  rq_init_comm_if_connected(9, "1")
  rq_init_comm_if_connected(2, "2")
  rq_init_comm_if_connected(3, "3")
  rq_init_comm_if_connected(4, "4")
  rq_print_connected_grippers()
  rq_gripper_communication_thread = run rq_gripper_communication()
  set_closed_norm(97.6470588235294, "1")
  set_open_norm(1.1764705882352942, "1")
  set_closed_mm(0.0, "1")
  set_open_mm(53.0, "1")
  set_closed_norm(100.0, "2")
  set_open_norm(0.0, "2")
  set_closed_mm(0.0, "2")
  set_open_mm(50.0, "2")
  set_closed_norm(100.0, "3")
  set_open_norm(0.0, "3")
  set_closed_mm(0.0, "3")
  set_open_mm(50.0, "3")
  set_closed_norm(100.0, "4")
  set_open_norm(0.0, "4")
  set_closed_mm(0.0, "4")
  set_open_mm(50.0, "4")
  rq_current_limit_enabled = False
  while(not rq_gripper_communication_thread_started):
      sleep(0.008)
  end
  # end: URCap Installation Node
  step_count_652fcfe5_f3e5_4323_a28e_c4dd7c99f65c = 0.0
  thread Step_Counter_Thread_2d5c0d0e_2884_4a5b_ab92_48b0595c18f1():
    while (True):
      step_count_652fcfe5_f3e5_4323_a28e_c4dd7c99f65c = step_count_652fcfe5_f3e5_4323_a28e_c4dd7c99f65c + 1.0
      sync()
    end
  end
  run Step_Counter_Thread_2d5c0d0e_2884_4a5b_ab92_48b0595c18f1()
  global AMR_Position=struct(position_identifier=0, x1=0, x2=0, y1=0, y2=0, theta1=0, theta2=0)
  $ 2 "BeforeStart"
  $ 3 "Manual"
  $ 4 "Home (Safe)"
  movej([-1.2291867130198177, -1.2978880085432127, -1.8023901537060905, -1.6126269993759976, 1.5736085024106596, 0.3398721000491988], a=1.3962634015954636, v=1.0471975511965976)
  $ 5 "STATE≔'state'"
  global STATE=request_integer_from_primary_client("state")
  $ 6 "If STATE≟6"
  if (STATE == 6):
    $ 7 "Action≔'what'"
    global Action=request_integer_from_primary_client("what")
    $ 8 "If Action≟52"
    if (Action == 52):
      $ 9 "AMR_PosTarget≔'target'"
      global AMR_PosTarget=request_integer_from_primary_client("target")
    end
  end
  $ 10 "Robot Program"
  $ 11 "PreSettings"
  $ 12 "AMR_TargetList≔[1,2,3,4,5,21,22,23,24,31,32,33,34,35,36,37,38,41]"
  global AMR_TargetList=[1,2,3,4,5,21,22,23,24,31,32,33,34,35,36,37,38,41]
  $ 13 "AMR_Done≔ False "
  global AMR_Done=  False
  $ 14 "AMR_PosActual≔T2O_Current_Pos"
  global AMR_PosActual=modbus_get_signal_status("T2O_Current_Pos")
  $ 15 "AMR_Attemps≔T2O_Nav_Attemps"
  global AMR_Attemps=modbus_get_signal_status("T2O_Nav_Attemps")
  $ 16 "AMR_Battery≔MiR_Battery_Lvl"
  global AMR_Battery=modbus_get_signal_status("MiR_Battery_Lvl")
  $ 17 "AMR_Charging≔(T2O_Charging≟1)"
  global AMR_Charging=(modbus_get_signal_status("T2O_Charging") == 1)
  $ 18 "AMR_Position≔struct(position_identifier=T2O_Current_Pos, x1=MiR_Position_X1, x2=MiR_Position_X2, y1=MiR_Position_Y1, y2=MiR_Position_Y2, theta1=MiR_Theta_1, theta2=MiR_Theta_2) "
  global AMR_Position=struct(position_identifier=modbus_get_signal_status("T2O_Current_Pos"), x1=modbus_get_signal_status("MiR_Position_X1"), x2=modbus_get_signal_status("MiR_Position_X2"), y1=modbus_get_signal_status("MiR_Position_Y1"), y2=modbus_get_signal_status("MiR_Position_Y2"), theta1=modbus_get_signal_status("MiR_Theta_1"), theta2=modbus_get_signal_status("MiR_Theta_2"))
  $ 19 "If MiR_Mode≠7"
  if (modbus_get_signal_status("MiR_Mode") != 7):
    $ 20 "Error"
    $ 21 "set_error(ERROR_AMR_WRONG_MODE)"
    set_error(ERROR_AMR_WRONG_MODE)
    $ 22 "AMR_Done≔ True "
    global AMR_Done=  True
  end
  $ 23 "'=========='"
  # '=========='
  $ 24 "Switch STATE"
  switch_1 = STATE
  $ 25 "Case 1"
  if (1 == switch_1):
    $ 26 "stopping"
    $ 27 "If T2O_Done≟1 and O2T_Acknowledge≟0"
    if (modbus_get_signal_status("T2O_Done") == 1  and  modbus_get_signal_status("O2T_Acknowledge") == 0):
      $ 28 "Set O2T_Acknowledge=1"
      modbus_set_output_register("O2T_Acknowledge", 1)
    end
    $ 29 "Set MiR_CMD_Stop=On"
    modbus_set_output_signal("MiR_CMD_Stop", True)
    $ 30 "If MiR_State≠3 and MiR_State≠5"
    if (modbus_get_signal_status("MiR_State") != 3  and  modbus_get_signal_status("MiR_State") != 5):
      $ 31 "AMR_Position.position_identifier = 0"
      AMR_Position.position_identifier = 0
      $ 32 "AMR_Done≔ True "
      global AMR_Done=  True
    end
  elif (2 == switch_1):
    $ 33 "Case 2"
    $ 34 "stopped"
    $ 35 "Set MiR_CMD_Stop=Off"
    modbus_set_output_signal("MiR_CMD_Stop", False)
  elif (3 == switch_1):
    $ 36 "Case 3"
    $ 37 "resetting"
    $ 38 "Set O2T_Mis_Main=Off"
    modbus_set_output_signal("O2T_Mis_Main", False)
    $ 39 "Set O2T_Mis_Charge=Off"
    modbus_set_output_signal("O2T_Mis_Charge", False)
    $ 40 "If MiR_Mis_Queue>0"
    if (modbus_get_signal_status("MiR_Mis_Queue")>0):
      $ 41 "Set MiR_CMD_Clear_Q=On"
      modbus_set_output_signal("MiR_CMD_Clear_Q", True)
      $ 42 "Wait MiR_Mis_Queue≟0"
      while (not(modbus_get_signal_status("MiR_Mis_Queue") == 0)):
        sync()
      end
      $ 43 "Set MiR_CMD_Clear_Q=Off"
      modbus_set_output_signal("MiR_CMD_Clear_Q", False)
    end
    $ 44 "If MiR_Error_ID≠0"
    if (modbus_get_signal_status("MiR_Error_ID") != 0):
      $ 45 "Set MiR_CMD_Clear_E=On"
      modbus_set_output_signal("MiR_CMD_Clear_E", True)
      $ 46 "Wait MiR_Error_ID≟0"
      while (not(modbus_get_signal_status("MiR_Error_ID") == 0)):
        sync()
      end
      $ 47 "Set MiR_CMD_Clear_E=Off"
      modbus_set_output_signal("MiR_CMD_Clear_E", False)
    end
    $ 48 "Set O2T_Action=0"
    modbus_set_output_register("O2T_Action", 0)
    $ 49 "Set O2T_Acknowledge=0"
    modbus_set_output_register("O2T_Acknowledge", 0)
    $ 50 "Set O2T_Target_Pos=0"
    modbus_set_output_register("O2T_Target_Pos", 0)
    $ 51 "Set O2T_Footprint=0"
    modbus_set_output_register("O2T_Footprint", 0)
    $ 52 "Set O2T_ProtectOff=0"
    modbus_set_output_register("O2T_ProtectOff", 0)
    $ 53 "Set O2T_Dock=0"
    modbus_set_output_register("O2T_Dock", 0)
    $ 54 "AMR_Attemps≔0"
    global AMR_Attemps=0
    $ 55 "AMR_PosTarget≔0"
    global AMR_PosTarget=0
    $ 56 "AMR_Step≔0"
    global AMR_Step=0
    $ 57 "AMR_AtTarget≔ False "
    global AMR_AtTarget=  False
    $ 58 "If MiR_State≟4 or MiR_State≟3 or MiR_State≟10"
    if (modbus_get_signal_status("MiR_State") == 4  or  modbus_get_signal_status("MiR_State") == 3  or  modbus_get_signal_status("MiR_State") == 10):
      $ 59 "AMR_Done≔ True "
      global AMR_Done=  True
    end
  elif (5 == switch_1):
    $ 60 "Case 5"
    $ 61 "starting"
    $ 62 "If MiR_State≟4"
    if (modbus_get_signal_status("MiR_State") == 4):
      $ 63 "Set MiR_CMD_Start=On"
      modbus_set_output_signal("MiR_CMD_Start", True)
      $ 64 "Wait MiR_State≠4"
      while (not(modbus_get_signal_status("MiR_State") != 4)):
        sync()
      end
      $ 65 "Set MiR_CMD_Start=Off"
      modbus_set_output_signal("MiR_CMD_Start", False)
      $ 66 "AMR_Done≔ True "
      global AMR_Done=  True
    else:
      $ 67 "ElseIf MiR_State≟10"
      if (modbus_get_signal_status("MiR_State") == 10):
        $ 68 "'MiR in protective stop. Wait'"
        # 'MiR in protective stop. Wait'
        $ 69 "AMR_Done≔ True "
        global AMR_Done=  True
      else:
        $ 70 "ElseIf MiR_State≟3"
        if (modbus_get_signal_status("MiR_State") == 3):
          $ 71 "AMR_Done≔ True "
          global AMR_Done=  True
        end
      end
    end
  elif (6 == switch_1):
    $ 72 "Case 6"
    $ 73 "execute"
    $ 74 "AMR_AtTarget≔(AMR_PosActual≟AMR_PosTarget)"
    global AMR_AtTarget=(AMR_PosActual == AMR_PosTarget)
    $ 75 "Switch AMR_Step"
    switch_2 = AMR_Step
    $ 76 "Case 0"
    if (0 == switch_2):
      $ 77 "If  not AMR_AtTarget"
      if (  not  AMR_AtTarget):
        $ 78 "AMR_Step≔1"
        global AMR_Step=1
      else:
        $ 79 "Else" "noBreak"
        $ 80 "AMR_Done≔ True "
        global AMR_Done=  True
      end
    elif (1 == switch_2):
      $ 81 "Case 1"
      $ 82 "general Settings"
      $ 83 "Set O2T_Acknowledge=0"
      modbus_set_output_register("O2T_Acknowledge", 0)
      $ 84 "check for error"
      $ 85 "If OBJ_Picked and MiR_State≟10"
      if (OBJ_Picked  and  modbus_get_signal_status("MiR_State") == 10):
        $ 86 "Error"
        $ 87 "set_error(ERROR_ROBOT_ARM_NOT_IN_HOME_POSE)"
        set_error(ERROR_ROBOT_ARM_NOT_IN_HOME_POSE)
        $ 88 "Action≔0"
        global Action=0
      else:
        $ 89 "ElseIf  not found_in_list(AMR_PosTarget, AMR_TargetList)"
        if (  not  found_in_list(AMR_PosTarget, AMR_TargetList)):
          $ 90 "Error"
          $ 91 "set_error(ERROR_UNKNOWN_POSE)"
          set_error(ERROR_UNKNOWN_POSE)
          $ 92 "Action≔0"
          global Action=0
        end
      end
      $ 93 "If MiR_State≟3"
      if (modbus_get_signal_status("MiR_State") == 3):
        $ 94 "Set MiR_CMD_Start=Off"
        modbus_set_output_signal("MiR_CMD_Start", False)
        $ 95 "Switch Action"
        switch_3 = Action
        $ 96 "Case 51"
        if (51 == switch_3):
          $ 97 "Charge"
          $ 98 "'trigger the charging mission'"
          # 'trigger the charging mission'
          $ 99 "'target pos is predefined'"
          # 'target pos is predefined'
          $ 100 "Set O2T_Footprint=0"
          modbus_set_output_register("O2T_Footprint", 0)
          $ 101 "Set O2T_Action=1"
          modbus_set_output_register("O2T_Action", 1)
        elif (52 == switch_3):
          $ 102 "Case 52"
          $ 103 "Navigate"
          $ 104 "'trigger the standard missoin'"
          # 'trigger the standard missoin'
          $ 105 "Set O2T_Footprint=AMR_FootprintID"
          modbus_set_output_register("O2T_Footprint", AMR_FootprintID)
          $ 106 "Set O2T_Target_Pos=AMR_PosTarget"
          modbus_set_output_register("O2T_Target_Pos", AMR_PosTarget)
          $ 107 "Set O2T_Action=2"
          modbus_set_output_register("O2T_Action", 2)
        end
        $ 108 "If MiR_Mis_Queue≟0"
        if (modbus_get_signal_status("MiR_Mis_Queue") == 0):
          $ 109 "Set O2T_Mis_Main=On"
          modbus_set_output_signal("O2T_Mis_Main", True)
          $ 110 "Wait MiR_Mis_Queue≥1"
          while (not(modbus_get_signal_status("MiR_Mis_Queue") >= 1)):
            sync()
          end
          $ 111 "Set O2T_Mis_Main=Off"
          modbus_set_output_signal("O2T_Mis_Main", False)
        end
      else:
        $ 112 "ElseIf MiR_State≟4"
        if (modbus_get_signal_status("MiR_State") == 4):
          $ 113 "Set MiR_CMD_Start=On"
          modbus_set_output_signal("MiR_CMD_Start", True)
        else:
          $ 114 "ElseIf MiR_State≟5"
          if (modbus_get_signal_status("MiR_State") == 5):
            $ 115 "AMR_Step≔2"
            global AMR_Step=2
          else:
            $ 116 "ElseIf MiR_State≟10"
            if (modbus_get_signal_status("MiR_State") == 10):
              $ 117 "'AMR still in safeguard stop'"
              # 'AMR still in safeguard stop'
            end
          end
        end
      end
    elif (2 == switch_2):
      $ 118 "Case 2"
      $ 119 "acknowledge handshake"
      $ 120 "If T2O_Done≟1 and O2T_Acknowledge≟0"
      if (modbus_get_signal_status("T2O_Done") == 1  and  modbus_get_signal_status("O2T_Acknowledge") == 0):
        $ 121 "Set O2T_Acknowledge=1"
        modbus_set_output_register("O2T_Acknowledge", 1)
      else:
        $ 122 "ElseIf T2O_Done≟0 and O2T_Acknowledge≟1"
        if (modbus_get_signal_status("T2O_Done") == 0  and  modbus_get_signal_status("O2T_Acknowledge") == 1):
          $ 123 "Set O2T_Acknowledge=0"
          modbus_set_output_register("O2T_Acknowledge", 0)
          $ 124 "AMR_AtTarget≔(AMR_PosActual≟AMR_PosTarget)"
          global AMR_AtTarget=(AMR_PosActual == AMR_PosTarget)
          $ 125 "AMR_Done≔ True "
          global AMR_Done=  True
        end
      end
    end
    $ 126 "translate errors"
    $ 127 "If AMR_Done"
    if (AMR_Done):
      $ 128 "Switch T2O_Error_ID"
      switch_2 = modbus_get_signal_status("T2O_Error_ID")
      $ 129 "Case 2003"
      if (2003 == switch_2):
        $ 130 "error"
        $ 131 "set_error(ERROR_NOT_DOCKED)"
        set_error(ERROR_NOT_DOCKED)
      elif (2007 == switch_2):
        $ 132 "Case 2007"
        $ 133 "error"
        $ 134 "set_error(ERROR_NOT_REACHABLE_TARGET)"
        set_error(ERROR_NOT_REACHABLE_TARGET)
      elif (2008 == switch_2):
        $ 135 "Case 2008"
        $ 136 "error"
        $ 137 "set_error(ERROR_CHARGING_NOT_STARTED)"
        set_error(ERROR_CHARGING_NOT_STARTED)
      end
    end
  elif (7 == switch_1):
    $ 138 "Case 7"
    $ 139 "completing"
    $ 140 "If MiR_Mis_Queue>0"
    if (modbus_get_signal_status("MiR_Mis_Queue")>0):
      $ 141 "Set MiR_CMD_Abort=On"
      modbus_set_output_signal("MiR_CMD_Abort", True)
      $ 142 "Wait MiR_Mis_Queue≟0"
      while (not(modbus_get_signal_status("MiR_Mis_Queue") == 0)):
        sync()
      end
      $ 143 "Set MiR_CMD_Abort=Off"
      modbus_set_output_signal("MiR_CMD_Abort", False)
    end
    $ 144 "If MiR_State≟3 or MiR_State≟10"
    if (modbus_get_signal_status("MiR_State") == 3  or  modbus_get_signal_status("MiR_State") == 10):
      $ 145 "AMR_Done≔ True "
      global AMR_Done=  True
    end
  elif (9 == switch_1):
    $ 146 "Case 9"
    $ 147 "holding"
    $ 148 "Set MiR_CMD_Abort=On"
    modbus_set_output_signal("MiR_CMD_Abort", True)
    $ 149 "If MiR_State≟3 or MiR_State≟10"
    if (modbus_get_signal_status("MiR_State") == 3  or  modbus_get_signal_status("MiR_State") == 10):
      $ 150 "Set MiR_CMD_Abort=Off"
      modbus_set_output_signal("MiR_CMD_Abort", False)
      $ 151 "AMR_Done≔ True "
      global AMR_Done=  True
    end
  elif (11 == switch_1):
    $ 152 "Case 11"
    $ 153 "unholding"
    $ 154 "Set MiR_CMD_Start=On"
    modbus_set_output_signal("MiR_CMD_Start", True)
    $ 155 "If MiR_State≠4"
    if (modbus_get_signal_status("MiR_State") != 4):
      $ 156 "Set MiR_CMD_Start=Off"
      modbus_set_output_signal("MiR_CMD_Start", False)
      $ 157 "AMR_Step≔0"
      global AMR_Step=0
      $ 158 "AMR_Done≔ True "
      global AMR_Done=  True
    end
  elif (12 == switch_1):
    $ 159 "Case 12"
    $ 160 "suspending"
    $ 161 "'none'"
    # 'none'
  elif (14 == switch_1):
    $ 162 "Case 14"
    $ 163 "unsuspending"
    $ 164 "'none'"
    # 'none'
  elif (15 == switch_1):
    $ 165 "Case 15"
    $ 166 "aborting"
    $ 167 "Set MiR_CMD_Abort=On"
    modbus_set_output_signal("MiR_CMD_Abort", True)
    $ 168 "Wait MiR_State≟3"
    while (not(modbus_get_signal_status("MiR_State") == 3)):
      sync()
    end
    $ 169 "Set MiR_CMD_Abort=Off"
    modbus_set_output_signal("MiR_CMD_Abort", False)
  elif (17 == switch_1):
    $ 170 "Case 17"
    $ 171 "clearing"
    $ 172 "If MiR_Error_ID≠0"
    if (modbus_get_signal_status("MiR_Error_ID") != 0):
      $ 173 "Set MiR_CMD_Clear_E=On"
      modbus_set_output_signal("MiR_CMD_Clear_E", True)
      $ 174 "Wait MiR_Error_ID≟0"
      while (not(modbus_get_signal_status("MiR_Error_ID") == 0)):
        sync()
      end
      $ 175 "Set MiR_CMD_Clear_E=Off"
      modbus_set_output_signal("MiR_CMD_Clear_E", False)
    end
    $ 176 "If MiR_Error_ID≟0"
    if (modbus_get_signal_status("MiR_Error_ID") == 0):
      $ 177 "AMR_Done≔ True "
      global AMR_Done=  True
    end
  end
  $ 178 "'=========='"
  # '=========='
  $ 179 "PostSettings"
  $ 180 "AMR_Position≔struct(position_identifier=T2O_Current_Pos, x1=MiR_Position_X1, x2=MiR_Position_X2, y1=MiR_Position_Y1, y2=MiR_Position_Y2, theta1=MiR_Theta_1, theta2=MiR_Theta_2) "
  global AMR_Position=struct(position_identifier=modbus_get_signal_status("T2O_Current_Pos"), x1=modbus_get_signal_status("MiR_Position_X1"), x2=modbus_get_signal_status("MiR_Position_X2"), y1=modbus_get_signal_status("MiR_Position_Y1"), y2=modbus_get_signal_status("MiR_Position_Y2"), theta1=modbus_get_signal_status("MiR_Theta_1"), theta2=modbus_get_signal_status("MiR_Theta_2"))
end
